(* IEC 61131-3 sources: llm-plc-st-eval/data/definitivo/gemini-3.1-pro-preview/I3/zero_shot, 3 files *)

(* ---- ejec_1.st ---- *)
```iecst
FUNCTION_BLOCK FB_Alarmas
VAR_INPUT
    alm1 : BOOL; // Causa de alarma 1 (Prioridad Alta)
    alm2 : BOOL; // Causa de alarma 2 (Prioridad Media)
    alm3 : BOOL; // Causa de alarma 3 (Prioridad Baja)
    ack1 : BOOL; // Reconocimiento alarma 1
    ack2 : BOOL; // Reconocimiento alarma 2
    ack3 : BOOL; // Reconocimiento alarma 3
END_VAR

VAR_OUTPUT
    sirena : BOOL;   // Sirena activa si hay alguna alarma presente
    codigoAlm : INT; // Código de la alarma de mayor prioridad (1, 2, 3 o 0)
END_VAR

VAR
    memAlm1 : BOOL; // Memoria de retención para alarma 1
    memAlm2 : BOOL; // Memoria de retención para alarma 2
    memAlm3 : BOOL; // Memoria de retención para alarma 3
END_VAR

// 1. Lógica de retención y reconocimiento de alarmas
// La alarma se activa si la causa está presente.
// Se mantiene retenida mientras no se reciba el 'ack' correspondiente.
// Si la causa sigue presente, el 'ack' no tiene efecto (almX fuerza el TRUE).
memAlm1 := alm1 OR (memAlm1 AND NOT ack1);
memAlm2 := alm2 OR (memAlm2 AND NOT ack2);
memAlm3 := alm3 OR (memAlm3 AND NOT ack3);

// 2. Lógica de activación de la sirena
// Se enciende si cualquiera de las alarmas retenidas está activa
sirena := memAlm1 OR memAlm2 OR memAlm3;

// 3. Lógica de prioridad para el código de alarma
// Se evalúa en orden descendente de prioridad (Alta -> Media -> Baja)
IF memAlm1 THEN
    codigoAlm := 1;
ELSIF memAlm2 THEN
    codigoAlm := 2;
ELSIF memAlm3 THEN
    codigoAlm := 3;
ELSE
    codigoAlm := 0; // Ninguna alarma activa
END_IF;

END_FUNCTION_BLOCK
```

(* ---- ejec_2.st ---- *)
```iecst
FUNCTION_BLOCK FB_Alarmas
VAR_INPUT
    alm1 : BOOL; // Causa de alarma 1 (Prioridad Alta)
    alm2 : BOOL; // Causa de alarma 2 (Prioridad Media)
    alm3 : BOOL; // Causa de alarma 3 (Prioridad Baja)
    ack1 : BOOL; // Reconocimiento alarma 1
    ack2 : BOOL; // Reconocimiento alarma 2
    ack3 : BOOL; // Reconocimiento alarma 3
END_VAR

VAR_OUTPUT
    sirena : BOOL;   // Sirena activa si hay alguna alarma presente
    codigoAlm : INT; // Código de alarma de mayor prioridad (1, 2, 3 o 0)
END_VAR

VAR
    memAlm1 : BOOL; // Memoria de retención alarma 1
    memAlm2 : BOOL; // Memoria de retención alarma 2
    memAlm3 : BOOL; // Memoria de retención alarma 3
END_VAR

// Gestión de retención y reconocimiento (Alarma 1)
// Se activa con la causa. El ACK solo funciona si la causa (alm1) ya desapareció.
IF alm1 THEN
    memAlm1 := TRUE;
ELSIF ack1 THEN
    memAlm1 := FALSE;
END_IF;

// Gestión de retención y reconocimiento (Alarma 2)
IF alm2 THEN
    memAlm2 := TRUE;
ELSIF ack2 THEN
    memAlm2 := FALSE;
END_IF;

// Gestión de retención y reconocimiento (Alarma 3)
IF alm3 THEN
    memAlm3 := TRUE;
ELSIF ack3 THEN
    memAlm3 := FALSE;
END_IF;

// Activación de la sirena (cualquier alarma retenida la enciende)
sirena := memAlm1 OR memAlm2 OR memAlm3;

// Evaluación de prioridad para el código de salida
IF memAlm1 THEN
    codigoAlm := 1; // Prioridad Alta
ELSIF memAlm2 THEN
    codigoAlm := 2; // Prioridad Media
ELSIF memAlm3 THEN
    codigoAlm := 3; // Prioridad Baja
ELSE
    codigoAlm := 0; // Sin alarmas
END_IF;

END_FUNCTION_BLOCK
```

(* ---- ejec_3.st ---- *)
```iecst
FUNCTION_BLOCK FB_Alarmas
VAR_INPUT
    alm1 : BOOL; // Causa alarma 1 (Prioridad Alta)
    alm2 : BOOL; // Causa alarma 2 (Prioridad Media)
    alm3 : BOOL; // Causa alarma 3 (Prioridad Baja)
    ack1 : BOOL; // Reconocimiento alarma 1
    ack2 : BOOL; // Reconocimiento alarma 2
    ack3 : BOOL; // Reconocimiento alarma 3
END_VAR

VAR_OUTPUT
    sirena : BOOL;   // Sirena activa si hay alguna alarma presente
    codigoAlm : INT; // Código de la alarma de mayor prioridad (1, 2, 3 o 0 si no hay)
END_VAR

VAR
    estadoAlm1 : BOOL; // Estado retenido de la alarma 1
    estadoAlm2 : BOOL; // Estado retenido de la alarma 2
    estadoAlm3 : BOOL; // Estado retenido de la alarma 3
END_VAR

// 1. Lógica de retención (latch) y reconocimiento
// La alarma se activa si la causa está presente.
// Se mantiene activa mientras no se reconozca (ack).
// Si la causa sigue presente, el ack no tiene efecto (almX domina).
estadoAlm1 := alm1 OR (estadoAlm1 AND NOT ack1);
estadoAlm2 := alm2 OR (estadoAlm2 AND NOT ack2);
estadoAlm3 := alm3 OR (estadoAlm3 AND NOT ack3);

// 2. Lógica de prioridad para el código de alarma
// Se evalúa en orden descendente de prioridad (1 -> 2 -> 3)
IF estadoAlm1 THEN
    codigoAlm := 1;
ELSIF estadoAlm2 THEN
    codigoAlm := 2;
ELSIF estadoAlm3 THEN
    codigoAlm := 3;
ELSE
    codigoAlm := 0;
END_IF;

// 3. Lógica de activación de la sirena
// Se enciende si cualquiera de los estados retenidos es verdadero
sirena := estadoAlm1 OR estadoAlm2 OR estadoAlm3;

END_FUNCTION_BLOCK
```
